// TIA Portal V21 export
// export: Created 2026-11-10T07:35:03.6323856Z, ExportSetting WithDefaults, DisplayName Totally Integrated Automation Portal, DisplayVersion V21 Update 3, DisplayName STEP 7 Professional, DisplayVersion V21 Update 3, DisplayName STEP 7 Safety, DisplayVersion V21, DisplayName Tech WebApplication, DisplayVersion V21, DisplayName WinCC Basic/Comfort/Advanced, DisplayVersion V21 Update 3, DisplayName WinCC Unified, DisplayVersion V21 Update 3
FUNCTION_BLOCK "FB_Lad_ex038"   // FB13, LAD
{ S7_Optimized_Access := 'TRUE' }
VERSION : 0.1
// stored: AutoNumber true, IsIECCheckEnabled false, IsRetainMemResEnabled false, MemoryReserve 100, SetENOAutomatically false, UDAEnableTagReadback false
   VAR_INPUT
      v_size : DInt;
   END_VAR
   VAR_OUTPUT
      v_out : WString;
   END_VAR
BEGIN

REGION Network 1: GetInstanceName - Read out name of the read instance
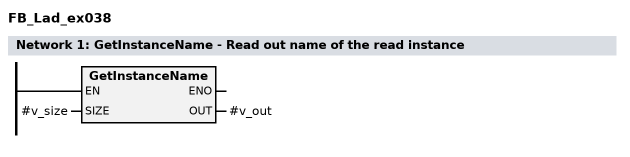
   RUNG wire#powerrail
      GetInstanceName(size := #v_size, OUT => #v_out)
   END_RUNG
   // the same network as SCL:
   GetInstanceName(size := #v_size, OUT => #v_out);
END_REGION
END_FUNCTION_BLOCK
